(* IEC 61131-3 sources: kns-pump-station/tests/POUs/Model/FB_PlantModel_Test, 41 files *)

(* ---- FB_PlantModel_Test.decl.st ---- *)
// Назначение: набор coUnit для FB_PlantModel (и FB_AnalogSensorSim, F_FloatContact, F_FaultInjEqual) — модель
//             объекта целиком: начальное состояние входов ПЛК, баланс массы, установившийся режим против эталона,
//             согласованность при разном шаге (ускорении), команды модели и сброс импульсов, ливень по команде,
//             отказы датчиков 4–20 мА, поплавки, вентилятор, инъекции насосов и счётчик их изменений, кнопки,
//             сухой ход и засор, осушенный приёмок, «время назад», время суток, предел шага. Время —
//             PL.FB_FakeTime; ожидаемые значения — эталон tools_project/plant_reference.py.
// Автор:      kr0nsch
// Версия:     0.1.0
// Документ:   docs/DESIGN.md, разделы 11.3, 14.1
FUNCTION_BLOCK FB_PlantModel_Test EXTENDS coUnit.FB_TestSuite
VAR CONSTANT
    T_STEP : TIME := T#1S;            // шаг модели в тесте (k = 50 при цикле 20 мс)
    T_FINE : TIME := T#100MS;         // мелкий шаг
    UI_FREF_50HZ : UINT := 5000;
    UI_FREF_87PCT : UINT := 4350;     // 43,5 Гц
    R_EPS_MA : REAL := 2.0E-3;        // допуск тока датчика, мА
    R_EPS_M : REAL := 1.0E-4;         // допуск уровня, м
    UI_FAULT_FIELDS : UDINT := 23;    // полей ST_FaultInjection в проверке счётчика
    T_SUBSTEP : TIME := T#200MS;      // шаг вызова = один подшаг SIM_DT_SUBSTEP
    R_INFLOW_EDGE_M3H : REAL := 2160.003;   // поднимает 0,29 м за 0,2 с до 0,3000000052 м
    DW_NAN : DWORD := 16#7FC00000;
END_VAR

(* ---- AiFaultCurrents.method.decl.st ---- *)
// Инъекции датчика LT101 (уровень 1,2 м, 7,84 мА): обрыв 0, FailLow 3,0, FailHigh 22, UnderRange 3,7,
// OverRange 20,8, Forced — заданный ток; Freeze держит ток при изменении уровня; индекс SIM_AI_PT201
// действует только на PT201.
METHOD PRIVATE AiFaultCurrents
VAR
    fbTime : PL.FB_FakeTime;    // подменное время
    fbDut : FB_PlantModel;      // проверяемая модель
    stCfg : ST_SimCfg;          // параметры по умолчанию
    stCmd : ST_SimCmd;          // команды модели
    stFault : ST_FaultInjection;  // инъекции
END_VAR

(* ---- AirLockAndClogCurrents.method.decl.st ---- *)
// Сухой ход Н1 на 100 %: подача 0, ток 10,75 А (регистр 108); засор Н2 на 100 %: подача 75,01 м³/ч,
// ток 34,30 А (регистр 343) — PMI-15. Уровень держится на 1,4 м (приток равен подаче).
METHOD PRIVATE AirLockAndClogCurrents
VAR
    fbTime : PL.FB_FakeTime;    // подменное время
    fbDut : FB_PlantModel;      // проверяемая модель
    stCfg : ST_SimCfg;          // параметры по умолчанию
    stCmd : ST_SimCmd;          // команды модели
    stFault : ST_FaultInjection;  // инъекции
    uiI : UINT;
END_VAR

(* ---- AirLockAndClogCurrents.method.impl.st ---- *)
coUnit.TEST('PlantModel_AirLockAndClogCurrents');

stCmd.xInflowOverride := TRUE;
stCmd.rInflowOverride_m3h := 75.012261;
stFault.axAirLock[1] := TRUE;
stFault.axClog[2] := TRUE;
fbDut.axRun[1] := TRUE;
fbDut.auiFref[1] := UI_FREF_50HZ;
fbDut.axRun[2] := TRUE;
fbDut.auiFref[2] := UI_FREF_50HZ;
fbDut(itfTime := fbTime, stCfg := stCfg, stCmd := stCmd, stFault := stFault);
FOR uiI := 1 TO 11 DO
    fbTime.Advance(tStep := T_STEP);
    fbDut(itfTime := fbTime, stCfg := stCfg, stCmd := stCmd, stFault := stFault);
END_FOR
stCmd.xSetLevel := TRUE;
stCmd.rSetLevel_m := 1.4;
FOR uiI := 1 TO 3 DO
    fbTime.Advance(tStep := T_STEP);
    fbDut(itfTime := fbTime, stCfg := stCfg, stCmd := stCmd, stFault := stFault);
END_FOR
// ref: hydraulic.air_lock_100, hydraulic.clog_100
AssertEquals_REAL(Expected := 0.0, Actual := fbDut.stSts.arPumpFlow_m3h[1], Delta := 0.0,
                  Message := 'air lock: no flow');
AssertEquals_REAL(Expected := 10.752, Actual := fbDut.stSts.arCurrent_A[1], Delta := 0.01,
                  Message := 'air lock current');
AssertEquals_UINT(Expected := 108, Actual := fbDut.stIo.uiIT111, Message := 'air lock register');
AssertEquals_REAL(Expected := 75.012261, Actual := fbDut.stSts.arPumpFlow_m3h[2], Delta := 0.05,
                  Message := 'clog flow');
AssertEquals_REAL(Expected := 34.299021, Actual := fbDut.stSts.arCurrent_A[2], Delta := 0.01,
                  Message := 'clog current');
AssertEquals_UINT(Expected := 343, Actual := fbDut.stIo.uiIT121, Message := 'clog register');

coUnit.TEST_FINISHED();

(* ---- ButtonsPulse.method.decl.st ---- *)
// xPressReset: HS501 нажата 500 мс (0,4 с — нажата, 0,5 с — отпущена), импульс команды сброшен; HS502 не нажата.
METHOD PRIVATE ButtonsPulse
VAR
    fbTime : PL.FB_FakeTime;    // подменное время
    fbDut : FB_PlantModel;      // проверяемая модель
    stCfg : ST_SimCfg;          // параметры по умолчанию
    stCmd : ST_SimCmd;          // команды модели
    stFault : ST_FaultInjection;  // инъекции
    uiI : UINT;
END_VAR

(* ---- ButtonsPulse.method.impl.st ---- *)
coUnit.TEST('PlantModel_ButtonsPulse');

stCmd.xPressReset := TRUE;
fbDut(itfTime := fbTime, stCfg := stCfg, stCmd := stCmd, stFault := stFault);
AssertFalse(Condition := stCmd.xPressReset, Message := 'pulse reset');
AssertTrue(Condition := fbDut.stIo.xHS501, Message := 'HS501 pressed');
AssertFalse(Condition := fbDut.stIo.xHS502, Message := 'HS502 not pressed');
FOR uiI := 1 TO 4 DO
    fbTime.Advance(tStep := T_FINE);
    fbDut(itfTime := fbTime, stCfg := stCfg, stCmd := stCmd, stFault := stFault);
END_FOR
AssertTrue(Condition := fbDut.stIo.xHS501, Message := 'HS501 pressed at 0.4 s');
FOR uiI := 1 TO 1 DO
    fbTime.Advance(tStep := T_FINE);
    fbDut(itfTime := fbTime, stCfg := stCfg, stCmd := stCmd, stFault := stFault);
END_FOR
AssertFalse(Condition := fbDut.stIo.xHS501, Message := 'HS501 released at 0.5 s');
stCmd.xPressSilence := TRUE;
fbDut(itfTime := fbTime, stCfg := stCfg, stCmd := stCmd, stFault := stFault);
AssertTrue(Condition := fbDut.stIo.xHS502 AND NOT stCmd.xPressSilence, Message := 'HS502 pressed');

coUnit.TEST_FINISHED();

(* ---- ClearFaultsZeroesFaultsOnly.method.decl.st ---- *)
// xClearFaults снимает все инъекции (значения по умолчанию типа: газы < 0 — фон) и сбрасывает импульс;
// приток, уровень и параметры не меняются.
METHOD PRIVATE ClearFaultsZeroesFaultsOnly
VAR
    fbTime : PL.FB_FakeTime;    // подменное время
    fbDut : FB_PlantModel;      // проверяемая модель
    stCfg : ST_SimCfg;          // параметры по умолчанию
    stCmd : ST_SimCmd;          // команды модели
    stFault : ST_FaultInjection;  // инъекции
    stNoFaults : ST_FaultInjection;  // значения по умолчанию
END_VAR

(* ---- DefaultsInitialState.method.decl.st ---- *)
// Первый вызов с параметрами по умолчанию: уровень 1,2 м (LT101 7,84 мА), насосы стоят (PT201 —
// столб 1,1772 бар = 5,8835 мА, FT202 4 мА), газы — фон (4,24 мА), поплавки и ввод в норме, ПЧ готовы
// (STW 16#0011), обмен исправен, TT403 18 °C, приток в 0 ч — 0,55 · 70 = 38,5 м³/ч.
METHOD PRIVATE DefaultsInitialState
VAR
    fbTime : PL.FB_FakeTime;    // подменное время
    fbDut : FB_PlantModel;      // проверяемая модель
    stCfg : ST_SimCfg;          // параметры по умолчанию
    stCmd : ST_SimCmd;          // команды модели
    stFault : ST_FaultInjection;  // инъекции
END_VAR

(* ---- FanNoFeedback.method.decl.st ---- *)
// В1: блок-контакт следует команде через 1 с (0,9 с — нет, 1,0 с — есть); xFanNoFeedback — ОС нет при
// поданной команде (V1.FTS, V1.FBL); xFanFault — V1_FLT; снятие команды — ОС пропадает через 1 с.
METHOD PRIVATE FanNoFeedback
VAR
    fbTime : PL.FB_FakeTime;    // подменное время
    fbDut : FB_PlantModel;      // проверяемая модель
    stCfg : ST_SimCfg;          // параметры по умолчанию
    stCmd : ST_SimCmd;          // команды модели
    stFault : ST_FaultInjection;  // инъекции
    uiI : UINT;
END_VAR

(* ---- FanNoFeedback.method.impl.st ---- *)
coUnit.TEST('PlantModel_FanNoFeedback');

fbDut.xV1Run := TRUE;
fbDut(itfTime := fbTime, stCfg := stCfg, stCmd := stCmd, stFault := stFault);
FOR uiI := 1 TO 9 DO
    fbTime.Advance(tStep := T_FINE);
    fbDut(itfTime := fbTime, stCfg := stCfg, stCmd := stCmd, stFault := stFault);
END_FOR
AssertFalse(Condition := fbDut.stIo.xV1_RFB, Message := 'no feedback at 0.9 s');
FOR uiI := 1 TO 1 DO
    fbTime.Advance(tStep := T_FINE);
    fbDut(itfTime := fbTime, stCfg := stCfg, stCmd := stCmd, stFault := stFault);
END_FOR
AssertTrue(Condition := fbDut.stIo.xV1_RFB, Message := 'feedback at 1.0 s');
stFault.xFanNoFeedback := TRUE;
FOR uiI := 1 TO 1 DO
    fbTime.Advance(tStep := T_FINE);
    fbDut(itfTime := fbTime, stCfg := stCfg, stCmd := stCmd, stFault := stFault);
END_FOR
AssertFalse(Condition := fbDut.stIo.xV1_RFB, Message := 'feedback injection: no feedback');
stFault.xFanNoFeedback := FALSE;
stFault.xFanFault := TRUE;
FOR uiI := 1 TO 1 DO
    fbTime.Advance(tStep := T_FINE);
    fbDut(itfTime := fbTime, stCfg := stCfg, stCmd := stCmd, stFault := stFault);
END_FOR
AssertTrue(Condition := fbDut.stIo.xV1_FLT AND fbDut.stIo.xV1_RFB, Message := 'fan fault contact');
fbDut.xV1Run := FALSE;
FOR uiI := 1 TO 10 DO
    fbTime.Advance(tStep := T_FINE);
    fbDut(itfTime := fbTime, stCfg := stCfg, stCmd := stCmd, stFault := stFault);
END_FOR
AssertTrue(Condition := fbDut.stIo.xV1_RFB, Message := 'feedback held 0.9 s after stop');
FOR uiI := 1 TO 1 DO
    fbTime.Advance(tStep := T_FINE);
    fbDut(itfTime := fbTime, stCfg := stCfg, stCmd := stCmd, stFault := stFault);
END_FOR
AssertFalse(Condition := fbDut.stIo.xV1_RFB, Message := 'feedback drops 1.0 s after stop');

coUnit.TEST_FINISHED();

(* ---- FaultSeqCountsChanges.method.decl.st ---- *)
// Каждое изменение любого поля ST_FaultInjection (23 поля по очереди) увеличивает udiFaultSeq на 1;
// вызов без изменений — нет; xClearFaults — ещё одно изменение.
METHOD PRIVATE FaultSeqCountsChanges
VAR
    fbTime : PL.FB_FakeTime;    // подменное время
    fbDut : FB_PlantModel;      // проверяемая модель
    stCfg : ST_SimCfg;          // параметры по умолчанию
    stCmd : ST_SimCmd;          // команды модели
    stFault : ST_FaultInjection;  // инъекции
END_VAR

(* ---- FloatStuckNormalTripped.method.decl.st ---- *)
// Поплавки НЗ: LS102 срабатывает при уровне ≥ 4,20 м (FALSE), LS103 — при ≤ 0,40 м; StuckNormal —
// не срабатывает (TRUE), StuckTripped — сработал при любом уровне (FALSE).
METHOD PRIVATE FloatStuckNormalTripped
VAR
    fbTime : PL.FB_FakeTime;    // подменное время
    fbDut : FB_PlantModel;      // проверяемая модель
    stCfg : ST_SimCfg;          // параметры по умолчанию
    stCmd : ST_SimCmd;          // команды модели
    stFault : ST_FaultInjection;  // инъекции
END_VAR

(* ---- IntakeDryStopsPumping.method.decl.st ---- *)
// Уровень 0,25 м ниже приёмка: насос на 100 % не откачивает, уровень не падает, ток холостого хода 10,75 А.
METHOD PRIVATE IntakeDryStopsPumping
VAR
    fbTime : PL.FB_FakeTime;    // подменное время
    fbDut : FB_PlantModel;      // проверяемая модель
    stCfg : ST_SimCfg;          // параметры по умолчанию
    stCmd : ST_SimCmd;          // команды модели
    stFault : ST_FaultInjection;  // инъекции
    uiI : UINT;
END_VAR

(* ---- IntakeDryStopsPumping.method.impl.st ---- *)
coUnit.TEST('PlantModel_IntakeDryStopsPumping');

stCmd.xInflowOverride := TRUE;
stCmd.rInflowOverride_m3h := 0.0;
stCmd.xSetLevel := TRUE;
stCmd.rSetLevel_m := 0.25;
fbDut.axRun[1] := TRUE;
fbDut.auiFref[1] := UI_FREF_50HZ;
fbDut(itfTime := fbTime, stCfg := stCfg, stCmd := stCmd, stFault := stFault);
FOR uiI := 1 TO 12 DO
    fbTime.Advance(tStep := T_STEP);
    fbDut(itfTime := fbTime, stCfg := stCfg, stCmd := stCmd, stFault := stFault);
END_FOR
// ref: hydraulic.intake_dry
AssertEquals_REAL(Expected := 0.0, Actual := fbDut.stSts.rOutflow_m3h, Delta := 0.0, Message := 'no pumping');
AssertEquals_REAL(Expected := 0.25, Actual := fbDut.stSts.rLevel_m, Delta := R_EPS_M, Message := 'level kept');
AssertEquals_REAL(Expected := 10.752, Actual := fbDut.stSts.arCurrent_A[1], Delta := 0.01,
                  Message := 'dry running current');

coUnit.TEST_FINISHED();

(* ---- IntakeEdgeOutflowMatchesTank.method.decl.st ---- *)
// Отметка приёмка (0,30 м): решение «приёмок осушен» для гидравлики и для резервуара — одно и то же
// (по уровню LREAL резервуара). Уровень 0,29 м, насос 1 на 50 Гц; за шаг 0,2 с приток 2160,003 м³/ч
// поднимает его до 0,3000000052 м — в LREAL ниже отметки, а в REAL (0,30000001) уже на ней. Подача
// насоса (FT202, rOutflow_m3h), которую резервуар не откачивает, нарушала бы баланс массы. Затем
// установка уровня 1,0 м (подача есть) и 0,25 м (подачи нет) — шагами по 0,2 с (один подшаг).
METHOD PRIVATE IntakeEdgeOutflowMatchesTank
VAR
    fbTime : PL.FB_FakeTime;    // подменное время
    fbDut : FB_PlantModel;      // проверяемая модель
    stCfg : ST_SimCfg;          // параметры по умолчанию
    stCmd : ST_SimCmd;          // команды модели
    stFault : ST_FaultInjection;  // инъекции
    uiI : UINT;
END_VAR

(* ---- IntakeEdgeOutflowMatchesTank.method.impl.st ---- *)
coUnit.TEST('PlantModel_IntakeEdgeOutflowMatchesTank');

stCmd.xInflowOverride := TRUE;
stCmd.rInflowOverride_m3h := 0.0;
stCmd.xSetLevel := TRUE;
stCmd.rSetLevel_m := 0.29;
fbDut.axRun[1] := TRUE;
fbDut.auiFref[1] := UI_FREF_50HZ;
fbDut(itfTime := fbTime, stCfg := stCfg, stCmd := stCmd, stFault := stFault);
FOR uiI := 1 TO 12 DO
    fbTime.Advance(tStep := T_STEP);
    fbDut(itfTime := fbTime, stCfg := stCfg, stCmd := stCmd, stFault := stFault);
END_FOR
AssertEquals_REAL(Expected := 50.0, Actual := fbDut.stSts.arFreq_Hz[1], Delta := 1.0E-3, Message := 'drive at 50 Hz');
stCmd.rInflowOverride_m3h := R_INFLOW_EDGE_M3H;
fbTime.Advance(tStep := T_SUBSTEP);
fbDut(itfTime := fbTime, stCfg := stCfg, stCmd := stCmd, stFault := stFault);
stCmd.rInflowOverride_m3h := 0.0;
fbTime.Advance(tStep := T_SUBSTEP);
fbDut(itfTime := fbTime, stCfg := stCfg, stCmd := stCmd, stFault := stFault);
AssertTrue(Condition := fbDut.stSts.rLevel_m >= GVL_Const.SIM_PUMP_INTAKE_M, Message := 'REAL level at intake mark');
AssertEquals_REAL(Expected := 0.0, Actual := fbDut.stSts.rOutflow_m3h, Delta := 0.0,
                  Message := 'tank not drained: no outflow reported');
AssertEquals_REAL(Expected := 4.0, Actual := fbDut.stIo.rFT202_mA, Delta := R_EPS_MA, Message := 'FT202 zero flow');
stCmd.xSetLevel := TRUE;
stCmd.rSetLevel_m := 1.0;
fbTime.Advance(tStep := T_SUBSTEP);
fbDut(itfTime := fbTime, stCfg := stCfg, stCmd := stCmd, stFault := stFault);
AssertTrue(Condition := fbDut.stSts.rOutflow_m3h > 100.0, Message := 'pumping at 1.0 m');
AssertTrue(Condition := fbDut.stSts.rLevel_m < 1.0, Message := 'level falls at 1.0 m');
stCmd.xSetLevel := TRUE;
stCmd.rSetLevel_m := 0.25;
fbTime.Advance(tStep := T_SUBSTEP);
fbDut(itfTime := fbTime, stCfg := stCfg, stCmd := stCmd, stFault := stFault);
AssertEquals_REAL(Expected := 0.0, Actual := fbDut.stSts.rOutflow_m3h, Delta := 0.0,
                  Message := 'set below intake: no outflow in the same call');
AssertEquals_REAL(Expected := 0.25, Actual := fbDut.stSts.rLevel_m, Delta := R_EPS_M, Message := 'level kept 0.25 m');

coUnit.TEST_FINISHED();

(* ---- MassBalanceNoPumps.method.decl.st ---- *)
// Постоянный приток 60 м³/ч без насосов 10 мин: уровень растёт на 60 · (1/6) / 12 = 0,8333 м.
METHOD PRIVATE MassBalanceNoPumps
VAR
    fbTime : PL.FB_FakeTime;    // подменное время
    fbDut : FB_PlantModel;      // проверяемая модель
    stCfg : ST_SimCfg;          // параметры по умолчанию
    stCmd : ST_SimCmd;          // команды модели
    stFault : ST_FaultInjection;  // инъекции
    uiI : UINT;
END_VAR

(* ---- MassBalanceNoPumps.method.impl.st ---- *)
coUnit.TEST('PlantModel_MassBalanceNoPumps');

stCmd.xInflowOverride := TRUE;
stCmd.rInflowOverride_m3h := 60.0;
fbDut(itfTime := fbTime, stCfg := stCfg, stCmd := stCmd, stFault := stFault);
FOR uiI := 1 TO 600 DO
    fbTime.Advance(tStep := T_STEP);
    fbDut(itfTime := fbTime, stCfg := stCfg, stCmd := stCmd, stFault := stFault);
END_FOR
// ref: tank.balance_60_10min.dlevel_m
AssertEquals_REAL(Expected := 2.033333, Actual := fbDut.stSts.rLevel_m, Delta := R_EPS_M,
                  Message := 'level after 10 min');
AssertEquals_REAL(Expected := 60.0, Actual := fbDut.stSts.rInflow_m3h, Delta := 0.0, Message := 'inflow');
AssertEquals_REAL(Expected := 0.0, Actual := fbDut.stSts.rOutflow_m3h, Delta := 0.0, Message := 'no outflow');
AssertEquals_LREAL(Expected := 600.0, Actual := fbDut.stSts.lrSimTime_s, Delta := LREAL#1.0E-6,
                   Message := 'model time');

coUnit.TEST_FINISHED();

(* ---- MassBalanceTwoPumps.method.decl.st ---- *)
// Баланс массы с двумя насосами на 50 Гц (приток 120 м³/ч, уровень от 2,0 м): за 60 с изменение уровня равно
// сумме (Qin − Qout) · dt / 3600 / S по показанной подаче станции; подача станции — сумма подач насосов (равные
// насосы делят её поровну), FT202 показывает подачу станции (4 + 16 · Q / 500 мА).
METHOD PRIVATE MassBalanceTwoPumps
VAR
    fbTime : PL.FB_FakeTime;    // подменное время
    fbDut : FB_PlantModel;      // проверяемая модель
    stCfg : ST_SimCfg;          // параметры по умолчанию
    stCmd : ST_SimCmd;          // команды модели
    stFault : ST_FaultInjection;  // инъекции
    uiI : UINT;
    lrLevel0_m : LREAL;         // уровень в начале учёта
    lrExpected_m : LREAL;       // уровень по балансу показанных потоков
END_VAR

(* ---- MassBalanceTwoPumps.method.impl.st ---- *)
coUnit.TEST('PlantModel_MassBalanceTwoPumps');

stCmd.xInflowOverride := TRUE;
stCmd.rInflowOverride_m3h := 120.0;
stCmd.xSetLevel := TRUE;
stCmd.rSetLevel_m := 2.0;
fbDut.axRun[1] := TRUE;
fbDut.auiFref[1] := UI_FREF_50HZ;
fbDut.axRun[2] := TRUE;
fbDut.auiFref[2] := UI_FREF_50HZ;
fbDut(itfTime := fbTime, stCfg := stCfg, stCmd := stCmd, stFault := stFault);
FOR uiI := 1 TO 12 DO
    fbTime.Advance(tStep := T_STEP);
    fbDut(itfTime := fbTime, stCfg := stCfg, stCmd := stCmd, stFault := stFault);
END_FOR
lrLevel0_m := REAL_TO_LREAL(fbDut.stSts.rLevel_m);
lrExpected_m := lrLevel0_m;
FOR uiI := 1 TO 60 DO
    fbTime.Advance(tStep := T_STEP);
    fbDut(itfTime := fbTime, stCfg := stCfg, stCmd := stCmd, stFault := stFault);
    lrExpected_m := lrExpected_m + REAL_TO_LREAL(fbDut.stSts.rInflow_m3h - fbDut.stSts.rOutflow_m3h)
                    * PL.F_TimeToSec(tIn := T_STEP) / REAL_TO_LREAL(GVL_Const.SIM_S_PER_H)
                    / REAL_TO_LREAL(stCfg.rTankArea_m2);
END_FOR
// AssertEquals_REAL пропускает NaN: конечность проверяется отдельно
AssertTrue(Condition := PL.F_IsFinite(rIn := fbDut.stSts.rLevel_m) AND PL.F_IsFinite(rIn := fbDut.stSts.rOutflow_m3h)
           AND PL.F_IsFinite(rIn := fbDut.stIo.rFT202_mA), Message := 'outputs finite');
AssertTrue(Condition := fbDut.stSts.rOutflow_m3h > 190.0, Message := 'two pumps deliver about 198 m3/h');
AssertEquals_REAL(Expected := fbDut.stSts.arPumpFlow_m3h[1] + fbDut.stSts.arPumpFlow_m3h[2],
                  Actual := fbDut.stSts.rOutflow_m3h, Delta := 1.0E-3, Message := 'station flow = sum of pumps');
AssertEquals_REAL(Expected := fbDut.stSts.arPumpFlow_m3h[1], Actual := fbDut.stSts.arPumpFlow_m3h[2],
                  Delta := 1.0E-3, Message := 'equal pumps share equally');
AssertEquals_LREAL(Expected := lrExpected_m, Actual := REAL_TO_LREAL(fbDut.stSts.rLevel_m), Delta := LREAL#1.0E-4,
                   Message := 'level follows reported inflow and outflow');
AssertTrue(Condition := lrLevel0_m - REAL_TO_LREAL(fbDut.stSts.rLevel_m) > LREAL#0.1, Message := 'level falls 0.1 m');
AssertEquals_REAL(Expected := PL.GVL_Const.MA_ZERO + PL.GVL_Const.MA_SPAN * fbDut.stSts.rOutflow_m3h
                              / GVL_Const.SIM_FT202_RANGE_M3H,
                  Actual := fbDut.stIo.rFT202_mA, Delta := R_EPS_MA, Message := 'FT202 shows station flow');

coUnit.TEST_FINISHED();

(* ---- NanInjectionCountedOnce.method.decl.st ---- *)
// Неконечное значение в поле REAL инъекций (запись NaN по OPC UA или сценарием) — одно изменение, а не
// изменение в каждом вызове: иначе udiFaultSeq рос бы 50 раз в секунду и событие 101021 затирало бы журнал
// на 200 записей за секунды. Возврат к конечному значению — тоже одно изменение.
METHOD PRIVATE NanInjectionCountedOnce
VAR
    fbTime : PL.FB_FakeTime;    // подменное время
    fbDut : FB_PlantModel;      // проверяемая модель
    stCfg : ST_SimCfg;          // параметры по умолчанию
    stCmd : ST_SimCmd;          // команды модели
    stFault : ST_FaultInjection;  // инъекции
    uBits : PL.U_RealBits;
    uiI : UINT;
END_VAR

(* ---- NanInjectionCountedOnce.method.impl.st ---- *)
coUnit.TEST('PlantModel_NanInjectionCountedOnce');

uBits.dwValue := DW_NAN;
fbDut(itfTime := fbTime, stCfg := stCfg, stCmd := stCmd, stFault := stFault);
stFault.arAiForced_mA[GVL_Const.SIM_AI_PT201] := uBits.rValue;
FOR uiI := 1 TO 3 DO
    fbTime.Advance(tStep := T_STEP);
    fbDut(itfTime := fbTime, stCfg := stCfg, stCmd := stCmd, stFault := stFault);
END_FOR
AssertEquals_UDINT(Expected := 1, Actual := fbDut.stSts.udiFaultSeq, Message := 'forced NaN counted once');
stFault.rH2S_mgm3 := uBits.rValue;
FOR uiI := 1 TO 3 DO
    fbTime.Advance(tStep := T_STEP);
    fbDut(itfTime := fbTime, stCfg := stCfg, stCmd := stCmd, stFault := stFault);
END_FOR
AssertEquals_UDINT(Expected := 2, Actual := fbDut.stSts.udiFaultSeq, Message := 'gas NaN counted once');
// неконечная концентрация — ток отказа снизу (M7), не NaN во входе ПЛК
AssertTrue(Condition := PL.F_IsFinite(rIn := fbDut.stIo.rAT401_mA), Message := 'AT401 current finite');
AssertEquals_REAL(Expected := GVL_Const.SIM_MA_FAIL_LOW, Actual := fbDut.stIo.rAT401_mA, Delta := 0.0,
                  Message := 'NaN gas -> fail-low current');
stFault.arAiForced_mA[GVL_Const.SIM_AI_PT201] := 4.0;
FOR uiI := 1 TO 3 DO
    fbTime.Advance(tStep := T_STEP);
    fbDut(itfTime := fbTime, stCfg := stCfg, stCmd := stCmd, stFault := stFault);
END_FOR
AssertEquals_UDINT(Expected := 3, Actual := fbDut.stSts.udiFaultSeq, Message := 'NaN to finite counted once');

coUnit.TEST_FINISHED();

(* ---- OverflowTimeResolvedBySubsteps.method.decl.st ---- *)
// Шаг вызова 2 с (SIM_DT_MAX) делится на подшаги SIM_DT_SUBSTEP = 200 мс: уровень 4,595949 м, приток 250 м³/ч
// без насосов — отметка 4,6 м достигается в конце 4-го подшага (0,8 с), перелив — 7 подшагов = 1,4 с → 1 с.
// Одним шагом 2 с перелив был бы 2 с, подшагами по 0,4 с — 1,6 с → 2 с.
METHOD PRIVATE OverflowTimeResolvedBySubsteps
VAR
    fbTime : PL.FB_FakeTime;    // подменное время
    fbDut : FB_PlantModel;      // проверяемая модель
    stCfg : ST_SimCfg;          // параметры по умолчанию
    stCmd : ST_SimCmd;          // команды модели
    stFault : ST_FaultInjection;  // инъекции
END_VAR

(* ---- PerPumpSignalsIsolated.method.decl.st ---- *)
// Каждый насос — свои входы ПЛК (имена GVL_IO у насосов разные, блоки в модели явные). Для насоса i:
// инъекции перегрева, протечки, «Местного», аварии ПЧ и потери связи меняют только TS1i2, MS1i3, HS1i4,
// P10i_FLT, P10i_FCODE и xMbOk_RS485_1_Si; в работе только насоса i частота, ток, реле «Работа» — только у него.
METHOD PRIVATE PerPumpSignalsIsolated
VAR
    fbTime : PL.FB_FakeTime;    // подменное время
    fbDut : FB_PlantModel;      // проверяемая модель
    stCfg : ST_SimCfg;          // параметры по умолчанию
    stCmd : ST_SimCmd;          // команды модели
    stFault : ST_FaultInjection;  // инъекции
    stFaultNone : ST_FaultInjection;  // все инъекции сняты
    uiPump : UINT;              // насос с инъекцией или в работе
    uiJ : UINT;                 // проверяемый насос
    uiI : UINT;
    axTs : ARRAY[1..GVL_Const.STN_PUMP_COUNT] OF BOOL;      // TS1n2 (НЗ: TRUE — норма)
    axMs : ARRAY[1..GVL_Const.STN_PUMP_COUNT] OF BOOL;      // MS1n3
    axHs : ARRAY[1..GVL_Const.STN_PUMP_COUNT] OF BOOL;      // HS1n4
    axFlt : ARRAY[1..GVL_Const.STN_PUMP_COUNT] OF BOOL;     // P10n_FLT
    axRfb : ARRAY[1..GVL_Const.STN_PUMP_COUNT] OF BOOL;     // P10n_RFB
    axMbOk : ARRAY[1..GVL_Const.STN_PUMP_COUNT] OF BOOL;    // xMbOk_RS485_1_Sn
    auiFact : ARRAY[1..GVL_Const.STN_PUMP_COUNT] OF UINT;   // P10n_FACT
    auiIt : ARRAY[1..GVL_Const.STN_PUMP_COUNT] OF UINT;     // IT1n1
    auiFcode : ARRAY[1..GVL_Const.STN_PUMP_COUNT] OF UINT;  // P10n_FCODE
END_VAR

(* ---- PerPumpSignalsIsolated.method.impl.st ---- *)
coUnit.TEST('PlantModel_PerPumpSignalsIsolated');

fbDut(itfTime := fbTime, stCfg := stCfg, stCmd := stCmd, stFault := stFault);
FOR uiPump := 1 TO GVL_Const.STN_PUMP_COUNT DO
    // 1. Перегрев, протечка, «Местное», потеря связи насоса uiPump
    stFault := stFaultNone;
    stFault.axOverheat[uiPump] := TRUE;
    stFault.axLeak[uiPump] := TRUE;
    stFault.axLocal[uiPump] := TRUE;
    stFault.axVfdCommLoss[uiPump] := TRUE;
    fbTime.Advance(tStep := T_STEP);
    fbDut(itfTime := fbTime, stCfg := stCfg, stCmd := stCmd, stFault := stFault);
    axTs[1] := fbDut.stIo.xTS112;
    axTs[2] := fbDut.stIo.xTS122;
    axTs[3] := fbDut.stIo.xTS132;
    axMs[1] := fbDut.stIo.xMS113;
    axMs[2] := fbDut.stIo.xMS123;
    axMs[3] := fbDut.stIo.xMS133;
    axHs[1] := fbDut.stIo.xHS114;
    axHs[2] := fbDut.stIo.xHS124;
    axHs[3] := fbDut.stIo.xHS134;
    axFlt[1] := fbDut.stIo.xP101_FLT;
    axFlt[2] := fbDut.stIo.xP102_FLT;
    axFlt[3] := fbDut.stIo.xP103_FLT;
    axMbOk[1] := fbDut.stIo.xMbOk_RS485_1_S1;
    axMbOk[2] := fbDut.stIo.xMbOk_RS485_1_S2;
    axMbOk[3] := fbDut.stIo.xMbOk_RS485_1_S3;
    FOR uiJ := 1 TO GVL_Const.STN_PUMP_COUNT DO
        AssertTrue(Condition := axTs[uiJ] = (uiJ <> uiPump), Message := 'TS1n2 of its own pump only');
        AssertTrue(Condition := axMs[uiJ] = (uiJ = uiPump), Message := 'MS1n3 of its own pump only');
        AssertTrue(Condition := axHs[uiJ] = (uiJ = uiPump), Message := 'HS1n4 of its own pump only');
        AssertTrue(Condition := axFlt[uiJ] = (uiJ = uiPump), Message := 'overheat trips its own drive only');
        AssertTrue(Condition := axMbOk[uiJ] = (uiJ <> uiPump), Message := 'comm loss of its own slave only');
    END_FOR
    // 2. Авария ПЧ насоса uiPump (сначала исходное состояние: перегрев снят, ПЧ готовы)
    stFault := stFaultNone;
    stCmd.xResetPlant := TRUE;
    fbTime.Advance(tStep := T_STEP);
    fbDut(itfTime := fbTime, stCfg := stCfg, stCmd := stCmd, stFault := stFault);
    stFault.axVfdFault[uiPump] := TRUE;
    fbTime.Advance(tStep := T_STEP);
    fbDut(itfTime := fbTime, stCfg := stCfg, stCmd := stCmd, stFault := stFault);
    axFlt[1] := fbDut.stIo.xP101_FLT;
    axFlt[2] := fbDut.stIo.xP102_FLT;
    axFlt[3] := fbDut.stIo.xP103_FLT;
    auiFcode[1] := fbDut.stIo.uiP101_FCODE;
    auiFcode[2] := fbDut.stIo.uiP102_FCODE;
    auiFcode[3] := fbDut.stIo.uiP103_FCODE;
    FOR uiJ := 1 TO GVL_Const.STN_PUMP_COUNT DO
        AssertTrue(Condition := axFlt[uiJ] = (uiJ = uiPump), Message := 'drive fault of its own pump only');
    END_FOR
    AssertEquals_UINT(Expected := GVL_Const.SIM_VFD_FCODE_EXT, Actual := auiFcode[uiPump],
                      Message := 'own fault code 11');
    // 3. В работе только насос uiPump: частота, ток, реле «Работа»
    stFault := stFaultNone;
    stCmd.xResetPlant := TRUE;
    fbDut.axRun[uiPump] := TRUE;
    fbDut.auiFref[uiPump] := UI_FREF_50HZ;
    FOR uiI := 1 TO 12 DO
        fbTime.Advance(tStep := T_STEP);
        fbDut(itfTime := fbTime, stCfg := stCfg, stCmd := stCmd, stFault := stFault);
    END_FOR
    axRfb[1] := fbDut.stIo.xP101_RFB;
    axRfb[2] := fbDut.stIo.xP102_RFB;
    axRfb[3] := fbDut.stIo.xP103_RFB;
    auiFact[1] := fbDut.stIo.uiP101_FACT;
    auiFact[2] := fbDut.stIo.uiP102_FACT;
    auiFact[3] := fbDut.stIo.uiP103_FACT;
    auiIt[1] := fbDut.stIo.uiIT111;
    auiIt[2] := fbDut.stIo.uiIT121;
    auiIt[3] := fbDut.stIo.uiIT131;
    FOR uiJ := 1 TO GVL_Const.STN_PUMP_COUNT DO
        AssertTrue(Condition := axRfb[uiJ] = (uiJ = uiPump), Message := 'run relay of its own pump only');
        AssertTrue(Condition := (auiFact[uiJ] = UI_FREF_50HZ) = (uiJ = uiPump) AND (auiFact[uiJ] = 0) = (uiJ <> uiPump),
                   Message := 'FACT of its own drive only');
        AssertTrue(Condition := (auiIt[uiJ] > 0) = (uiJ = uiPump), Message := 'current register of its own drive only');
    END_FOR
    fbDut.axRun[uiPump] := FALSE;
    FOR uiI := 1 TO 12 DO
        fbTime.Advance(tStep := T_STEP);
        fbDut(itfTime := fbTime, stCfg := stCfg, stCmd := stCmd, stFault := stFault);
    END_FOR
END_FOR

coUnit.TEST_FINISHED();

(* ---- PumpAndStationInjectionsReachIo.method.decl.st ---- *)
// Инъекции доходят до входов ПЛК: авария ПЧ Н2 (FLT, STW.2, код 11), перегрев Н1 (TS112 = FALSE, авария
// ПЧ, код 12), протечка Н3, «Местное» Н2, потеря связи с ПЧ Н3, затопление, пожар, ИБП, дверь, газы,
// потеря связи с TT403 (значение замирает), пропадание напряжения (ES301, YS302, ПЧ без связи).
METHOD PRIVATE PumpAndStationInjectionsReachIo
VAR
    fbTime : PL.FB_FakeTime;    // подменное время
    fbDut : FB_PlantModel;      // проверяемая модель
    stCfg : ST_SimCfg;          // параметры по умолчанию
    stCmd : ST_SimCmd;          // команды модели
    stFault : ST_FaultInjection;  // инъекции
END_VAR

(* ---- ResetPlantClearsOverflowTime.method.decl.st ---- *)
// И0 (06 §5.2) перед каждой проверкой — xResetPlant: время перелива udiOverflow_s прошлой проверки
// обнуляется, иначе «перелива нет (SimSts.udiOverflow_s = 0)» PMI-20 и PMI-24 зависело бы от порядка
// проверок. Перелив: 4,55 м, приток 250 м³/ч без насосов, 60 с.
METHOD PRIVATE ResetPlantClearsOverflowTime
VAR
    fbTime : PL.FB_FakeTime;    // подменное время
    fbDut : FB_PlantModel;      // проверяемая модель
    stCfg : ST_SimCfg;          // параметры по умолчанию
    stCmd : ST_SimCmd;          // команды модели
    stFault : ST_FaultInjection;  // инъекции
    uiI : UINT;
END_VAR

(* ---- ResetPlantClearsOverflowTime.method.impl.st ---- *)
coUnit.TEST('PlantModel_ResetPlantClearsOverflowTime');

stCmd.xInflowOverride := TRUE;
stCmd.rInflowOverride_m3h := 250.0;
stCmd.xSetLevel := TRUE;
stCmd.rSetLevel_m := 4.55;
fbDut(itfTime := fbTime, stCfg := stCfg, stCmd := stCmd, stFault := stFault);
FOR uiI := 1 TO 60 DO
    fbTime.Advance(tStep := T_STEP);
    fbDut(itfTime := fbTime, stCfg := stCfg, stCmd := stCmd, stFault := stFault);
END_FOR
AssertTrue(Condition := fbDut.stSts.udiOverflow_s > 0, Message := 'overflow counted');
stCmd.rInflowOverride_m3h := 0.0;
stCmd.xResetPlant := TRUE;
fbTime.Advance(tStep := T_STEP);
fbDut(itfTime := fbTime, stCfg := stCfg, stCmd := stCmd, stFault := stFault);
AssertEquals_REAL(Expected := 1.2, Actual := fbDut.stSts.rLevel_m, Delta := R_EPS_M, Message := 'level 1.2 m');
AssertEquals_UDINT(Expected := 0, Actual := fbDut.stSts.udiOverflow_s, Message := 'overflow time cleared');

coUnit.TEST_FINISHED();

(* ---- ResetPlantRestoresLevelAndDrives.method.decl.st ---- *)
// И0 (06 §5.2): xClearFaults и xResetPlant в одном вызове — уровень 1,2 м, авария ПЧ снята без фронта
// CTW.2, ПЧ готов; пуск по проводу удержан — насос снова разгоняется.
METHOD PRIVATE ResetPlantRestoresLevelAndDrives
VAR
    fbTime : PL.FB_FakeTime;    // подменное время
    fbDut : FB_PlantModel;      // проверяемая модель
    stCfg : ST_SimCfg;          // параметры по умолчанию
    stCmd : ST_SimCmd;          // команды модели
    stFault : ST_FaultInjection;  // инъекции
    uiI : UINT;
END_VAR

(* ---- ResetPlantRestoresLevelAndDrives.method.impl.st ---- *)
coUnit.TEST('PlantModel_ResetPlantRestoresLevelAndDrives');

fbDut.axRun[1] := TRUE;
fbDut.auiFref[1] := UI_FREF_50HZ;
fbDut(itfTime := fbTime, stCfg := stCfg, stCmd := stCmd, stFault := stFault);
FOR uiI := 1 TO 3 DO
    fbTime.Advance(tStep := T_STEP);
    fbDut(itfTime := fbTime, stCfg := stCfg, stCmd := stCmd, stFault := stFault);
END_FOR
stCmd.xSetLevel := TRUE;
stCmd.rSetLevel_m := 3.0;
stFault.axVfdFault[1] := TRUE;
FOR uiI := 1 TO 1 DO
    fbTime.Advance(tStep := T_STEP);
    fbDut(itfTime := fbTime, stCfg := stCfg, stCmd := stCmd, stFault := stFault);
END_FOR
AssertTrue(Condition := fbDut.stIo.xP101_FLT, Message := 'drive faulted');
AssertEquals_REAL(Expected := 3.0, Actual := fbDut.stSts.rLevel_m, Delta := 0.01, Message := 'level 3 m');
stCmd.xClearFaults := TRUE;
stCmd.xResetPlant := TRUE;
FOR uiI := 1 TO 1 DO
    fbTime.Advance(tStep := T_STEP);
    fbDut(itfTime := fbTime, stCfg := stCfg, stCmd := stCmd, stFault := stFault);
END_FOR
AssertFalse(Condition := stCmd.xResetPlant OR stCmd.xClearFaults, Message := 'pulses reset');
AssertEquals_REAL(Expected := 1.2, Actual := fbDut.stSts.rLevel_m, Delta := 0.01, Message := 'level back to 1.2 m');
AssertFalse(Condition := fbDut.stIo.xP101_FLT, Message := 'drive fault cleared');
AssertTrue(Condition := (fbDut.stIo.wP101_STW AND GVL_Const.VFD_STW_READY) <> 0, Message := 'drive ready');
FOR uiI := 1 TO 1 DO
    fbTime.Advance(tStep := T_STEP);
    fbDut(itfTime := fbTime, stCfg := stCfg, stCmd := stCmd, stFault := stFault);
END_FOR
AssertTrue(Condition := fbDut.stSts.arFreq_Hz[1] > 0.0, Message := 'wired run restarts the pump');

coUnit.TEST_FINISHED();

(* ---- SetTimeOfDayKeepsDay.method.decl.st ---- *)
// xSetTimeOfDay 23,99 ч, через 60 с — сутки 1, 0,0067 ч; снова 8,0 ч — сутки 1 остаются, приток
// по профилю 112 м³/ч (ливни выключены).
METHOD PRIVATE SetTimeOfDayKeepsDay
VAR
    fbTime : PL.FB_FakeTime;    // подменное время
    fbDut : FB_PlantModel;      // проверяемая модель
    stCfg : ST_SimCfg;          // параметры по умолчанию
    stCmd : ST_SimCmd;          // команды модели
    stFault : ST_FaultInjection;  // инъекции
    uiI : UINT;
END_VAR

(* ---- SetTimeOfDayKeepsDay.method.impl.st ---- *)
coUnit.TEST('PlantModel_SetTimeOfDayKeepsDay');

stCfg.uiStormsPerDayMax := 0;
stCmd.xSetTimeOfDay := TRUE;
stCmd.rTimeOfDay_h := 23.99;
fbDut(itfTime := fbTime, stCfg := stCfg, stCmd := stCmd, stFault := stFault);
AssertFalse(Condition := stCmd.xSetTimeOfDay, Message := 'pulse reset');
AssertEquals_REAL(Expected := 23.99, Actual := fbDut.stSts.rTimeOfDay_h, Delta := 1.0E-4, Message := 'time of day set');
AssertEquals_UDINT(Expected := 0, Actual := fbDut.stSts.udiDay, Message := 'day 0');
FOR uiI := 1 TO 60 DO
    fbTime.Advance(tStep := T_STEP);
    fbDut(itfTime := fbTime, stCfg := stCfg, stCmd := stCmd, stFault := stFault);
END_FOR
AssertEquals_UDINT(Expected := 1, Actual := fbDut.stSts.udiDay, Message := 'next day after midnight');
AssertEquals_REAL(Expected := 0.006667, Actual := fbDut.stSts.rTimeOfDay_h, Delta := 1.0E-4, Message := '00:00:24');
stCmd.xSetTimeOfDay := TRUE;
stCmd.rTimeOfDay_h := 8.0;
fbDut(itfTime := fbTime, stCfg := stCfg, stCmd := stCmd, stFault := stFault);
AssertEquals_UDINT(Expected := 1, Actual := fbDut.stSts.udiDay, Message := 'day kept');
AssertEquals_REAL(Expected := 8.0, Actual := fbDut.stSts.rTimeOfDay_h, Delta := 1.0E-4, Message := '08:00');
// ref: inflow.profile.at_08h_m3h
AssertEquals_REAL(Expected := 112.0, Actual := fbDut.stSts.rInflow_m3h, Delta := 1.0E-3,
                  Message := 'profile inflow 112');

coUnit.TEST_FINISHED();

(* ---- SteadyStateOnePump87.method.decl.st ---- *)
// Один насос на 87 % (43,5 Гц), приток 120 м³/ч, уровень равновесия 1,23735 м (эталон): за 10 мин
// уровень не уходит, подача 120 м³/ч, PT201 6,9232 мА (1,8270 бар), FT202 7,84 мА, ток 19,29 А (193).
METHOD PRIVATE SteadyStateOnePump87
VAR
    fbTime : PL.FB_FakeTime;    // подменное время
    fbDut : FB_PlantModel;      // проверяемая модель
    stCfg : ST_SimCfg;          // параметры по умолчанию
    stCmd : ST_SimCmd;          // команды модели
    stFault : ST_FaultInjection;  // инъекции
    uiI : UINT;
END_VAR

(* ---- SteadyStateOnePump87.method.impl.st ---- *)
coUnit.TEST('PlantModel_SteadyStateOnePump87');

stCmd.xInflowOverride := TRUE;
stCmd.rInflowOverride_m3h := 120.0;
fbDut.axRun[1] := TRUE;
fbDut.auiFref[1] := UI_FREF_87PCT;
fbDut(itfTime := fbTime, stCfg := stCfg, stCmd := stCmd, stFault := stFault);
FOR uiI := 1 TO 15 DO
    fbTime.Advance(tStep := T_STEP);
    fbDut(itfTime := fbTime, stCfg := stCfg, stCmd := stCmd, stFault := stFault);
END_FOR
// ref: steady.one_pump_87_inflow_120.level_m
stCmd.xSetLevel := TRUE;
stCmd.rSetLevel_m := 1.23735;
FOR uiI := 1 TO 600 DO
    fbTime.Advance(tStep := T_STEP);
    fbDut(itfTime := fbTime, stCfg := stCfg, stCmd := stCmd, stFault := stFault);
END_FOR
AssertEquals_REAL(Expected := 43.5, Actual := fbDut.stSts.arFreq_Hz[1], Delta := 1.0E-3, Message := 'drive at 43.5 Hz');
// AssertEquals_REAL пропускает NaN: конечность проверяется отдельно
AssertTrue(Condition := PL.F_IsFinite(rIn := fbDut.stSts.rLevel_m) AND PL.F_IsFinite(rIn := fbDut.stSts.rOutflow_m3h)
           AND PL.F_IsFinite(rIn := fbDut.stIo.rPT201_mA) AND PL.F_IsFinite(rIn := fbDut.stSts.arCurrent_A[1]),
           Message := 'outputs finite');
// ref: steady.one_pump_87_inflow_120.*
AssertEquals_REAL(Expected := 1.23735, Actual := fbDut.stSts.rLevel_m, Delta := 2.0E-3,
                  Message := 'equilibrium level kept');
AssertEquals_REAL(Expected := 120.0, Actual := fbDut.stSts.rOutflow_m3h, Delta := 0.05, Message := 'outflow = inflow');
AssertEquals_REAL(Expected := 6.923223, Actual := fbDut.stIo.rPT201_mA, Delta := R_EPS_MA, Message := 'PT201 mA');
AssertEquals_REAL(Expected := 7.84, Actual := fbDut.stIo.rFT202_mA, Delta := R_EPS_MA, Message := 'FT202 mA');
AssertEquals_REAL(Expected := 19.290206, Actual := fbDut.stSts.arCurrent_A[1], Delta := 0.01,
                  Message := 'motor current');
AssertTrue(Condition := fbDut.stIo.uiIT111 >= 192 AND fbDut.stIo.uiIT111 <= 194, Message := 'current register 193');
AssertTrue(Condition := fbDut.stIo.xP101_RFB, Message := 'run relay');

coUnit.TEST_FINISHED();

(* ---- StepCappedAtMax.method.decl.st ---- *)
// Шаг часов 10 с за вызов (пауза задачи) обрезается до SIM_DT_MAX = 2 с времени модели.
METHOD PRIVATE StepCappedAtMax
VAR
    fbTime : PL.FB_FakeTime;    // подменное время
    fbDut : FB_PlantModel;      // проверяемая модель
    stCfg : ST_SimCfg;          // параметры по умолчанию
    stCmd : ST_SimCmd;          // команды модели
    stFault : ST_FaultInjection;  // инъекции
END_VAR

(* ---- StormNowTrapezoid.method.decl.st ---- *)
// xStormNow: трапеция 10 мин, пик 200 м³/ч (ливни генератора и профиль выключены): 45 с — 100,
// 90 с — 200, 300 с — 200, 495 с — 100, после 600 с — 0, ливень закончился. При постоянном притоке команда
// не действует, импульс сбрасывается.
METHOD PRIVATE StormNowTrapezoid
VAR
    fbTime : PL.FB_FakeTime;    // подменное время
    fbDut : FB_PlantModel;      // проверяемая модель
    stCfg : ST_SimCfg;          // параметры по умолчанию
    stCmd : ST_SimCmd;          // команды модели
    stFault : ST_FaultInjection;  // инъекции
    uiI : UINT;
END_VAR

(* ---- StormNowTrapezoid.method.impl.st ---- *)
coUnit.TEST('PlantModel_StormNowTrapezoid');

stCfg.uiStormsPerDayMax := 0;
stCfg.rInflowAvg_m3h := 0.0;
stCmd.xStormNow := TRUE;
stCmd.rStormPeak_m3h := 200.0;
stCmd.tStormDuration := T#10M;
fbDut(itfTime := fbTime, stCfg := stCfg, stCmd := stCmd, stFault := stFault);
AssertFalse(Condition := stCmd.xStormNow, Message := 'pulse reset');
AssertTrue(Condition := fbDut.stSts.xStormActive, Message := 'storm started');
FOR uiI := 1 TO 45 DO
    fbTime.Advance(tStep := T_STEP);
    fbDut(itfTime := fbTime, stCfg := stCfg, stCmd := stCmd, stFault := stFault);
END_FOR
AssertEquals_REAL(Expected := 100.0, Actual := fbDut.stSts.rStormInflow_m3h, Delta := 0.01, Message := 'half of rise');
AssertEquals_REAL(Expected := 100.0, Actual := fbDut.stSts.rInflow_m3h, Delta := 0.01, Message := 'inflow = storm');
FOR uiI := 1 TO 45 DO
    fbTime.Advance(tStep := T_STEP);
    fbDut(itfTime := fbTime, stCfg := stCfg, stCmd := stCmd, stFault := stFault);
END_FOR
AssertEquals_REAL(Expected := 200.0, Actual := fbDut.stSts.rStormInflow_m3h, Delta := 0.01, Message := 'end of rise');
FOR uiI := 1 TO 210 DO
    fbTime.Advance(tStep := T_STEP);
    fbDut(itfTime := fbTime, stCfg := stCfg, stCmd := stCmd, stFault := stFault);
END_FOR
AssertEquals_REAL(Expected := 200.0, Actual := fbDut.stSts.rStormInflow_m3h, Delta := 0.01, Message := 'plateau');
FOR uiI := 1 TO 195 DO
    fbTime.Advance(tStep := T_STEP);
    fbDut(itfTime := fbTime, stCfg := stCfg, stCmd := stCmd, stFault := stFault);
END_FOR
AssertEquals_REAL(Expected := 100.0, Actual := fbDut.stSts.rStormInflow_m3h, Delta := 0.01, Message := 'half of fall');
FOR uiI := 1 TO 106 DO
    fbTime.Advance(tStep := T_STEP);
    fbDut(itfTime := fbTime, stCfg := stCfg, stCmd := stCmd, stFault := stFault);
END_FOR
AssertEquals_REAL(Expected := 0.0, Actual := fbDut.stSts.rStormInflow_m3h, Delta := 0.0, Message := 'storm over');
AssertFalse(Condition := fbDut.stSts.xStormActive, Message := 'storm ended');
stCmd.xInflowOverride := TRUE;
stCmd.xStormNow := TRUE;
FOR uiI := 1 TO 1 DO
    fbTime.Advance(tStep := T_STEP);
    fbDut(itfTime := fbTime, stCfg := stCfg, stCmd := stCmd, stFault := stFault);
END_FOR
AssertFalse(Condition := stCmd.xStormNow OR fbDut.stSts.xStormActive, Message := 'ignored with inflow override');

coUnit.TEST_FINISHED();

(* ---- TimeAccelerationConsistency.method.decl.st ---- *)
// Одинаковый процесс (приток 100 м³/ч, насос 1 пущен на 50 Гц) шагом 100 мс (k = 5) и шагом 1 с (k = 50)
// за 60 с времени модели: одно время модели, частота 50 Гц, уровни расходятся меньше 5 мм (разница — только
// дискретность рампы ПЧ в шаге вызова; резервуар интегрируется подшагами ≤ 200 мс).
METHOD PRIVATE TimeAccelerationConsistency
VAR
    fbTimeA : PL.FB_FakeTime;
    fbTimeB : PL.FB_FakeTime;
    fbA : FB_PlantModel;        // шаг 100 мс
    fbB : FB_PlantModel;        // шаг 1 с
    stCfg : ST_SimCfg;
    stCmdA : ST_SimCmd;
    stCmdB : ST_SimCmd;
    stFaultA : ST_FaultInjection;
    stFaultB : ST_FaultInjection;
    uiI : UINT;
END_VAR

(* ---- TimeAccelerationConsistency.method.impl.st ---- *)
coUnit.TEST('PlantModel_TimeAccelerationConsistency');

stCmdA.xInflowOverride := TRUE;
stCmdA.rInflowOverride_m3h := 100.0;
stCmdB := stCmdA;
fbA.axRun[1] := TRUE;
fbA.auiFref[1] := UI_FREF_50HZ;
fbB.axRun[1] := TRUE;
fbB.auiFref[1] := UI_FREF_50HZ;
fbA(itfTime := fbTimeA, stCfg := stCfg, stCmd := stCmdA, stFault := stFaultA);
fbB(itfTime := fbTimeB, stCfg := stCfg, stCmd := stCmdB, stFault := stFaultB);
FOR uiI := 1 TO 600 DO
    fbTimeA.Advance(tStep := T_FINE);
    fbA(itfTime := fbTimeA, stCfg := stCfg, stCmd := stCmdA, stFault := stFaultA);
END_FOR
FOR uiI := 1 TO 60 DO
    fbTimeB.Advance(tStep := T_STEP);
    fbB(itfTime := fbTimeB, stCfg := stCfg, stCmd := stCmdB, stFault := stFaultB);
END_FOR
// AssertEquals_REAL пропускает NaN: конечность проверяется отдельно
AssertTrue(Condition := PL.F_IsFinite(rIn := fbA.stSts.rLevel_m) AND PL.F_IsFinite(rIn := fbB.stSts.rLevel_m)
           AND PL.F_IsFinite(rIn := fbA.stSts.rOutflow_m3h) AND PL.F_IsFinite(rIn := fbB.stSts.rOutflow_m3h),
           Message := 'outputs finite');
AssertEquals_LREAL(Expected := fbA.stSts.lrSimTime_s, Actual := fbB.stSts.lrSimTime_s, Delta := LREAL#1.0E-6,
                   Message := 'same model time');
AssertEquals_REAL(Expected := 50.0, Actual := fbA.stSts.arFreq_Hz[1], Delta := 1.0E-3, Message := 'A at 50 Hz');
AssertEquals_REAL(Expected := 50.0, Actual := fbB.stSts.arFreq_Hz[1], Delta := 1.0E-3, Message := 'B at 50 Hz');
AssertEquals_REAL(Expected := fbA.stSts.rLevel_m, Actual := fbB.stSts.rLevel_m, Delta := 5.0E-3,
                  Message := 'levels agree within 5 mm');
AssertEquals_REAL(Expected := fbA.stSts.rOutflow_m3h, Actual := fbB.stSts.rOutflow_m3h, Delta := 0.5,
                  Message := 'outflows agree');
AssertTrue(Condition := fbA.stSts.rLevel_m < 1.2, Message := 'pump outpaces inflow');

coUnit.TEST_FINISHED();

(* ---- TimeBackwardsHoldsState.method.decl.st ---- *)
// «Время назад»: шаг 0 — уровень и время модели не меняются; дальше модель продолжает.
METHOD PRIVATE TimeBackwardsHoldsState
VAR
    fbTime : PL.FB_FakeTime;    // подменное время
    fbDut : FB_PlantModel;      // проверяемая модель
    stCfg : ST_SimCfg;          // параметры по умолчанию
    stCmd : ST_SimCmd;          // команды модели
    stFault : ST_FaultInjection;  // инъекции
    uiI : UINT;
    rLevel : REAL;             // уровень до скачка времени
END_VAR

(* ---- TimeBackwardsHoldsState.method.impl.st ---- *)
coUnit.TEST('PlantModel_TimeBackwardsHoldsState');

stCmd.xInflowOverride := TRUE;
stCmd.rInflowOverride_m3h := 60.0;
fbDut(itfTime := fbTime, stCfg := stCfg, stCmd := stCmd, stFault := stFault);
FOR uiI := 1 TO 10 DO
    fbTime.Advance(tStep := T_STEP);
    fbDut(itfTime := fbTime, stCfg := stCfg, stCmd := stCmd, stFault := stFault);
END_FOR
rLevel := fbDut.stSts.rLevel_m;
fbTime.SetNow(ltValue := fbTime.Now() - LTIME#5S);
fbDut(itfTime := fbTime, stCfg := stCfg, stCmd := stCmd, stFault := stFault);
AssertEquals_REAL(Expected := rLevel, Actual := fbDut.stSts.rLevel_m, Delta := 0.0, Message := 'level held');
AssertEquals_LREAL(Expected := 10.0, Actual := fbDut.stSts.lrSimTime_s, Delta := LREAL#1.0E-9,
                   Message := 'model time held');
FOR uiI := 1 TO 1 DO
    fbTime.Advance(tStep := T_STEP);
    fbDut(itfTime := fbTime, stCfg := stCfg, stCmd := stCmd, stFault := stFault);
END_FOR
AssertEquals_LREAL(Expected := 11.0, Actual := fbDut.stSts.lrSimTime_s, Delta := LREAL#1.0E-9,
                   Message := 'model resumes');
AssertTrue(Condition := fbDut.stSts.rLevel_m > rLevel, Message := 'level rises again');

coUnit.TEST_FINISHED();
